SUBAPPLICATION Uebung_252_AX (* Section-Switcher BIT wie 251, lang: I1/I8 alle aus, I2/I7 alle ein, Start alle aus *)
  (* Standard: 61499-2; Description: Copyright (c) 2026 Meisterschulen am Ostbahnhof This program and the accompanying materials are made available under the terms of the Eclipse Public License 2.0 which is available at https://www.eclipse.org/legal/epl-2.0/ SPDX-License-Identifier: EPL-2.0 *)
  (* Version 1.0, 2026-11-05, Franz Höpfinger, Meisterschulen am Ostbahnhof, initial API and implementation and/or initial documentation *)
  PACKAGE Uebungen;
  IMPORT logiBUS::io::DI::logiBUS_DI::Input_I1;
  IMPORT logiBUS::io::DI::logiBUS_DI::Input_I2;
  IMPORT logiBUS::io::DI::logiBUS_DI::Input_I7;
  IMPORT logiBUS::io::DI::logiBUS_DI::Input_I8;
  IMPORT logiBUS::io::DI::logiBUS_DI_Events::BUTTON_SINGLE_CLICK;
  IMPORT logiBUS::io::DI::logiBUS_DI_Events::BUTTON_LONG_PRESS_START;
  IMPORT logiBUS::io::DQ::logiBUS_DO::Output_Q1;
  IMPORT logiBUS::io::DQ::logiBUS_DO::Output_Q2;
  IMPORT logiBUS::io::DQ::logiBUS_DO::Output_Q3;
  IMPORT logiBUS::io::DQ::logiBUS_DO::Output_Q4;
  IMPORT logiBUS::io::DQ::logiBUS_DO::Output_Q5;
  IMPORT logiBUS::io::DQ::logiBUS_DO::Output_Q6;
  IMPORT logiBUS::io::DQ::logiBUS_DO::Output_Q7;
  IMPORT logiBUS::io::DQ::logiBUS_DO::Output_Q8;
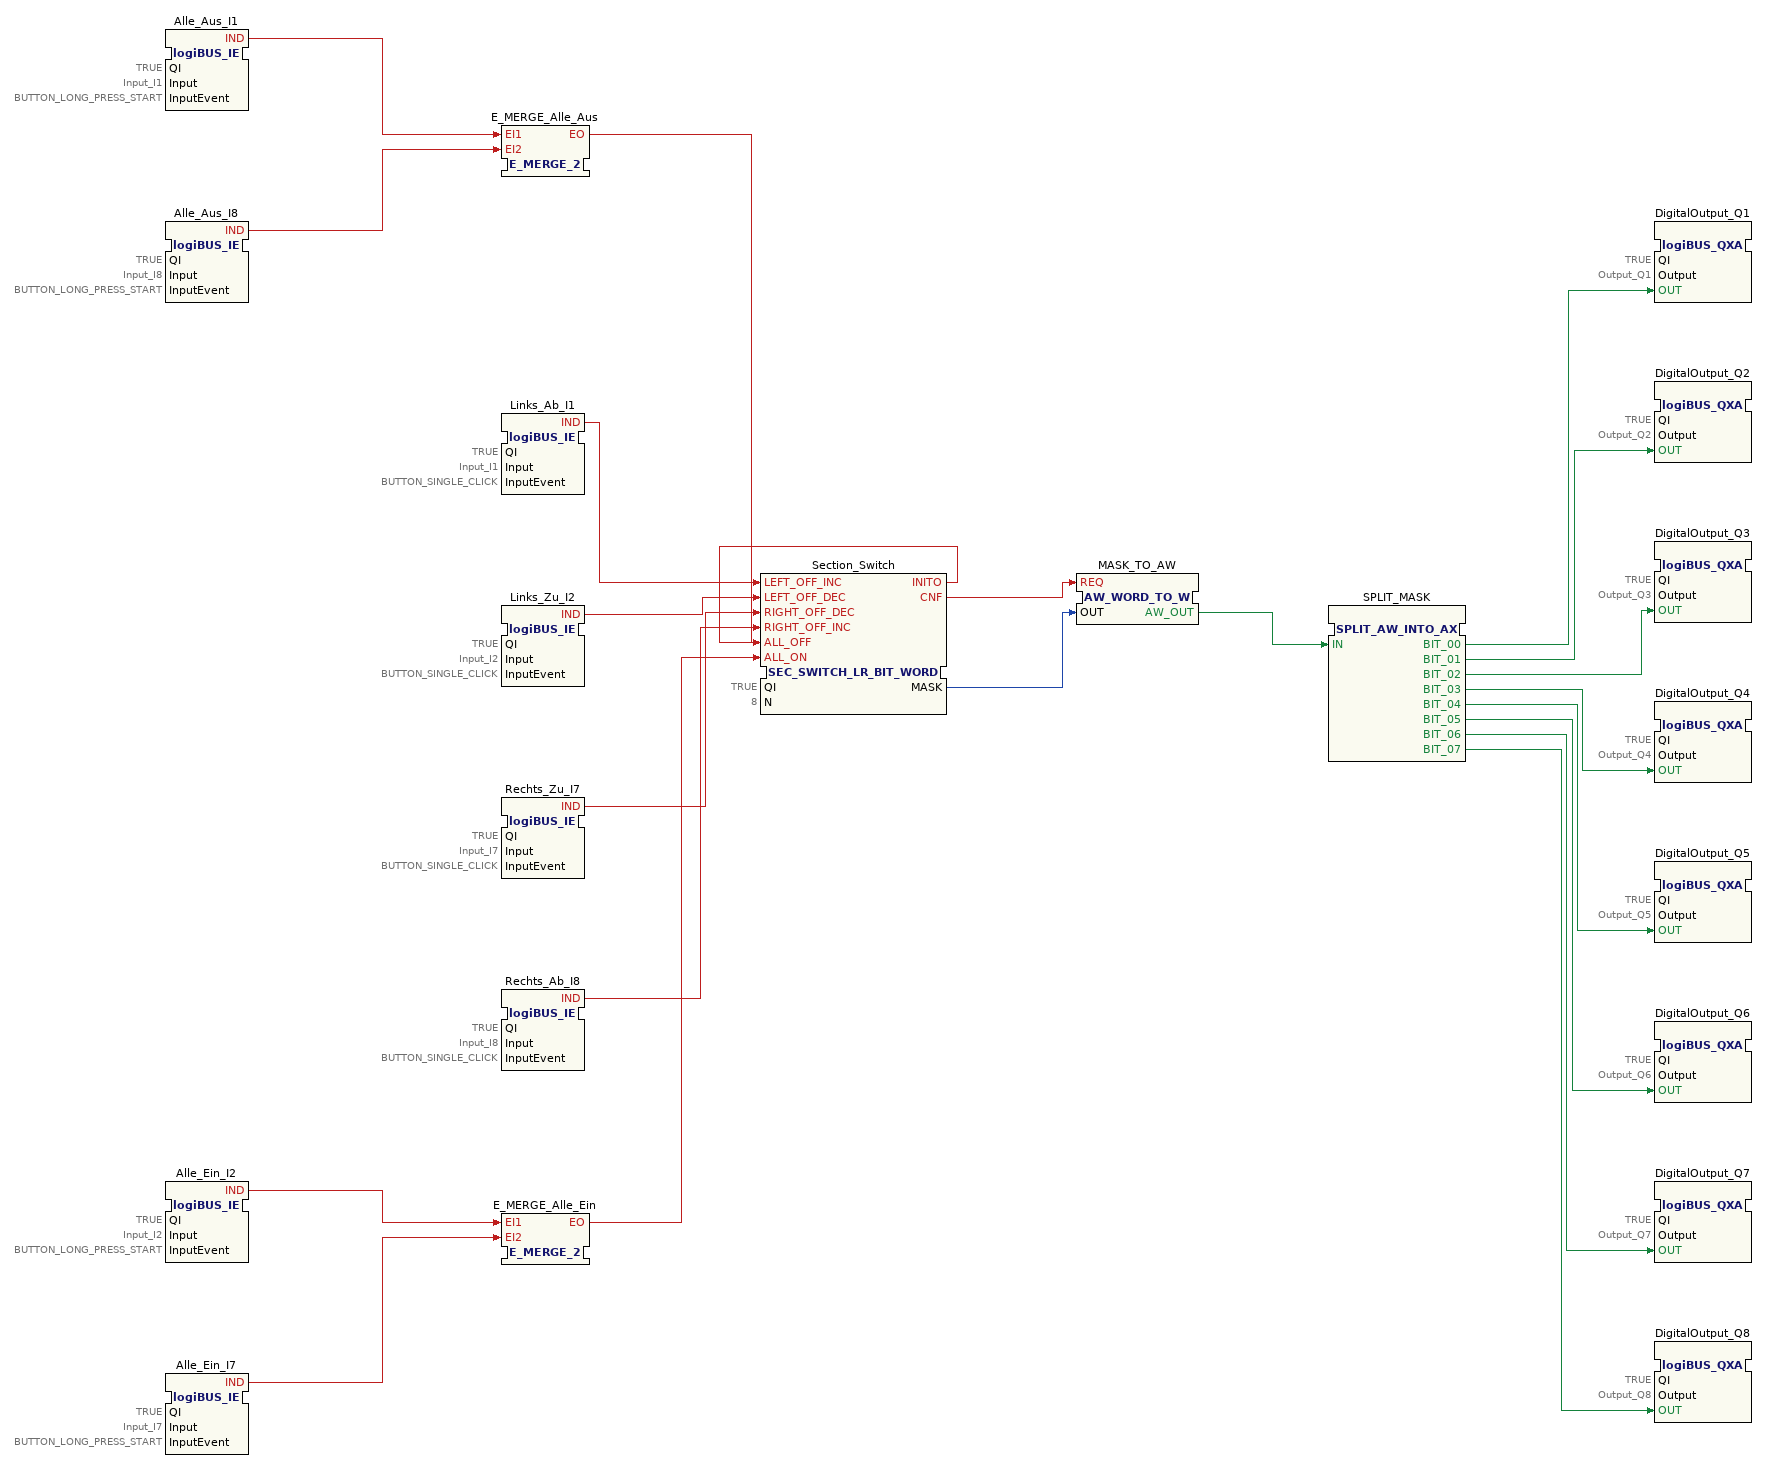
  FBS
    Links_Ab_I1 : logiBUS::io::DI::logiBUS_IE(QI := TRUE, Input := Input_I1, InputEvent := BUTTON_SINGLE_CLICK);
    Links_Zu_I2 : logiBUS::io::DI::logiBUS_IE(QI := TRUE, Input := Input_I2, InputEvent := BUTTON_SINGLE_CLICK);
    Rechts_Zu_I7 : logiBUS::io::DI::logiBUS_IE(QI := TRUE, Input := Input_I7, InputEvent := BUTTON_SINGLE_CLICK);
    Rechts_Ab_I8 : logiBUS::io::DI::logiBUS_IE(QI := TRUE, Input := Input_I8, InputEvent := BUTTON_SINGLE_CLICK);
    Section_Switch : logiBUS::sections::SEC_SWITCH_LR_BIT_WORD(QI := TRUE, N := 8); (* Startet sicher: INITO auf ALL_OFF, alle Sections aus *)
    MASK_TO_AW : adapter::conversion::unidirectional::AW_WORD_TO_W;
    SPLIT_MASK : adapter::splitting::SPLIT_AW_INTO_AX;
    DigitalOutput_Q1 : logiBUS::io::DQ::logiBUS_QXA(QI := TRUE, Output := Output_Q1);
    DigitalOutput_Q2 : logiBUS::io::DQ::logiBUS_QXA(QI := TRUE, Output := Output_Q2);
    DigitalOutput_Q3 : logiBUS::io::DQ::logiBUS_QXA(QI := TRUE, Output := Output_Q3);
    DigitalOutput_Q4 : logiBUS::io::DQ::logiBUS_QXA(QI := TRUE, Output := Output_Q4);
    DigitalOutput_Q5 : logiBUS::io::DQ::logiBUS_QXA(QI := TRUE, Output := Output_Q5);
    DigitalOutput_Q6 : logiBUS::io::DQ::logiBUS_QXA(QI := TRUE, Output := Output_Q6);
    DigitalOutput_Q7 : logiBUS::io::DQ::logiBUS_QXA(QI := TRUE, Output := Output_Q7);
    DigitalOutput_Q8 : logiBUS::io::DQ::logiBUS_QXA(QI := TRUE, Output := Output_Q8);
    Alle_Aus_I1 : logiBUS::io::DI::logiBUS_IE(QI := TRUE, Input := Input_I1, InputEvent := BUTTON_LONG_PRESS_START);
    Alle_Aus_I8 : logiBUS::io::DI::logiBUS_IE(QI := TRUE, Input := Input_I8, InputEvent := BUTTON_LONG_PRESS_START);
    Alle_Ein_I2 : logiBUS::io::DI::logiBUS_IE(QI := TRUE, Input := Input_I2, InputEvent := BUTTON_LONG_PRESS_START);
    Alle_Ein_I7 : logiBUS::io::DI::logiBUS_IE(QI := TRUE, Input := Input_I7, InputEvent := BUTTON_LONG_PRESS_START);
    E_MERGE_Alle_Aus : iec61499::events::E_MERGE_2;
    E_MERGE_Alle_Ein : iec61499::events::E_MERGE_2;
  END_FBS
  EVENT_CONNECTIONS
    Links_Ab_I1.IND TO Section_Switch.LEFT_OFF_INC;
    Links_Zu_I2.IND TO Section_Switch.LEFT_OFF_DEC;
    Rechts_Zu_I7.IND TO Section_Switch.RIGHT_OFF_DEC;
    Rechts_Ab_I8.IND TO Section_Switch.RIGHT_OFF_INC;
    Section_Switch.INITO TO Section_Switch.ALL_OFF;
    Section_Switch.CNF TO MASK_TO_AW.REQ;
    Alle_Aus_I1.IND TO E_MERGE_Alle_Aus.EI1;
    Alle_Aus_I8.IND TO E_MERGE_Alle_Aus.EI2;
    Alle_Ein_I2.IND TO E_MERGE_Alle_Ein.EI1;
    Alle_Ein_I7.IND TO E_MERGE_Alle_Ein.EI2;
    E_MERGE_Alle_Aus.EO TO Section_Switch.ALL_OFF;
    E_MERGE_Alle_Ein.EO TO Section_Switch.ALL_ON;
  END_CONNECTIONS
  DATA_CONNECTIONS
    Section_Switch.MASK TO MASK_TO_AW.OUT;
  END_CONNECTIONS
  ADAPTER_CONNECTIONS
    MASK_TO_AW.AW_OUT TO SPLIT_MASK.IN;
    SPLIT_MASK.BIT_00 TO DigitalOutput_Q1.OUT;
    SPLIT_MASK.BIT_01 TO DigitalOutput_Q2.OUT;
    SPLIT_MASK.BIT_02 TO DigitalOutput_Q3.OUT;
    SPLIT_MASK.BIT_03 TO DigitalOutput_Q4.OUT;
    SPLIT_MASK.BIT_04 TO DigitalOutput_Q5.OUT;
    SPLIT_MASK.BIT_05 TO DigitalOutput_Q6.OUT;
    SPLIT_MASK.BIT_06 TO DigitalOutput_Q7.OUT;
    SPLIT_MASK.BIT_07 TO DigitalOutput_Q8.OUT;
  END_CONNECTIONS
END_SUBAPPLICATION
